(* IEC 61131-3 sources: plc-iiot-stack/src/POUs/Iiot/F_IiotCmdResultText, 2 files *)

(* ---- F_IiotCmdResultText.decl.st ---- *)
// Назначение: имя E_CmdResult устройства для поля cmd_result (коды 1..9); прочие — пусто.
// Автор:      kr0nsch
// Версия:     0.1.0
// Документ:   docs/plc_mqtt.md, раздел «Команды»
FUNCTION F_IiotCmdResultText : STRING(GVL_Const.IIOT_TEXT_LEN)
VAR_INPUT
    iResult : INT;    // TO_INT(stSts.stCommon.eCmdResult)
END_VAR

(* ---- F_IiotCmdResultText.impl.st ---- *)
CASE iResult OF
    1:
        F_IiotCmdResultText := 'Accepted';
    2:
        F_IiotCmdResultText := 'RejectedMode';
    3:
        F_IiotCmdResultText := 'RejectedInterlock';
    4:
        F_IiotCmdResultText := 'RejectedPermit';
    5:
        F_IiotCmdResultText := 'RejectedInhibit';
    6:
        F_IiotCmdResultText := 'RejectedFault';
    7:
        F_IiotCmdResultText := 'RejectedState';
    8:
        F_IiotCmdResultText := 'RejectedNotSupported';
    9:
        F_IiotCmdResultText := 'RejectedCfg';
ELSE
    F_IiotCmdResultText := '';
END_CASE
